Fanuc KAREL source: kf00088.KL

-- PROVISIONAL review KL for V1013-1; original PC SHA256 c6c1aa35e554087b4ffd925d04ee35aea90e018146117ea2371e98504644338a
-- Incomplete behavior may be omitted. Consult companion uncertainty JSON. Do not deploy.
PROGRAM KF00088
%NOLOCKGROUP
BEGIN
  -- UNRESOLVED_PC offsets 5-28; opcodes 27,22,1C,31,4A
  -- UNRESOLVED_PC offsets 33-37; opcodes 7F
END KF00088
